// TIA Portal V18 export
DATA_BLOCK "DB_VFD_Data"   // DB8
{ S7_Optimized_Access := 'FALSE' }
   VAR
      ReadRegs : Array[0..18] of Word;
      forward : Bool;
      revers : Bool;
      stop : Bool;
      setFrequency : Real;   // 0020h - 40033
      outputFrequency : Real;   // 0021h - 40034 actual
      outputCurrent : Real;   // 0022h - 40035
      outputVoltage : Real;   // 0025h - 40038
      voltageZPT : Int;   // 0026h - 40039
      statusInputTerminals : Int;   // 0029h - 40042
      commands : Int;   // 0000h - 40001
      settingFrequency : Int;   // 0001h - 40002
      lastAlarm : Word;
      secondAlarm : Word;
      thirdAlarm : Word;
      alarms : Array[0..18] of Bool;
   END_VAR
BEGIN
END_DATA_BLOCK
